// The MONET telescope (FB_MonetTelescopeControl) on mock axes, scanned in the MONETS MAIN order (telescope first, then
// the axes). One Scan() is one PLC scan. The scenario tests own one rig each (VAR_INST of the test method) and call Scan()
// once per PLC cycle: the astronomical clock needs a real NT_GetTime round trip (up to about 5 s) before the telescope
// accepts a goto/slew/track, so a rig is not usable before ClockValid. Everything else counts scans, not time.
// Plan: BROTLib specs/plans/2026-10-21-telescope-state-machine-unification.md (D1, step 1).
{attribute 'enable_dynamic_creation'}
FUNCTION_BLOCK FB_MonetRig
VAR
	fbComm			: FB_LogRecordingComm;	// #287: the log of the rig can be watched (fbComm.sWatch, nWatchHits)
	fbElev			: FB_ElevationMock(comm := fbComm);
	fbAzim			: FB_AzimuthMock(comm := fbComm);
	fbDero			: FB_DerotatorMock(comm := fbComm);
	fbFocus			: FB_FocusMock(comm := fbComm);
	fbCovers		: FB_CoversMock(comm := fbComm);	// a HalfBROT.FB_CoverControl subclass, its FB_Init takes comm
	stCoverOut		: HalfBROT.ST_CoverOut;	// the process outputs of the covers and the focus block (HalfBROT 0.14.0: VAR_IN_OUT stOut); the mocks do not use them
	stFocusOut		: HalfBROT.ST_FocusOut;
	fbBrakeHyd		: FB_BrakeHydraulicsMock;
	fbPointing		: FB_PointingModelForward(AOFF := 0.0, BNP := 0.0, AN_A := 0.0, AE_A := 0.0, NPAE := 0.0, EOFF := 0.0, AN_E := 0.0, AE_E := 0.0, TF := 0.0);	// zero coefficients
	fbPointingInv	: FB_PointingModelInversion(fbPointing := fbPointing);
	fbTel			: FB_MonetTelescopeControl(comm := fbComm);
	fbWatchdog		: FB_MonetMqttWatchdog(comm := fbComm);	// for MonetSafeState_Tests (a method VAR_INST cannot refer to a sibling in its init list)
	nScans			: UDINT;
	bManual			: BOOL;	// MAIN calls SuspendAutomatic instead of the body while the cabinet selector is on manual
	nTimeDivisor	: UDINT := 1;	// the time seam of the telescope under test (SetTimeDivisor)
	bEstopIn		: BOOL;	// SafetyHandling.estop
	bSafetyIn		: BOOL;	// SafetyHandling.error
	bMainReadyIn	: BOOL := TRUE;	// PowerMonitoring.phaseOK (MAIN: bMainReady := ready)
	stMotion		: BROTLib.ST_MotionConfig;	// stMotion of the telescope under test (SetMotion), default = the struct defaults (#24 step 2c)
	fElevationMoveVelocityIn	: LREAL := 5.0;	// the deprecated alias input (SetElevationMoveVelocity), default = its old default; MONETS MAIN passes 3.0
END_VAR
VAR CONSTANT
	telescopeConfig	: ST_TelescopeConfig := (longitude := 20.810808, latitude := -32.375823, altitude := 1798.0,
											 azimuthPark := 175, elevationPark := 60, derotatorPark := 0, focusPark := 36.0,
											 azimuthHome := 175, elevationHome := 40, derotatorHome := 0,
											 name := 'MONET/S', diameter := 1.2, cabinet := 'Beckhoff', manufacturer := 'test',
											 mountOptions := 'ALT-AZ', mount := 'ALT_AZ');
END_VAR

// scans a homing takes on the three mock axes (default 3): a test that wants to act while the axes are homing makes it longer
METHOD SetHomeScans
VAR_INPUT
	nScans	: UINT;
END_VAR
fbElev.nMockHomeScans := nScans;
fbAzim.nMockHomeScans := nScans;
fbDero.nMockHomeScans := nScans;
END_METHOD

// scans a move takes on the three mock axes (default 60)
METHOD SetMoveScans
VAR_INPUT
	nScans	: UINT;
END_VAR
fbElev.nMockMoveScans := nScans;
fbAzim.nMockMoveScans := nScans;
fbDero.nMockMoveScans := nScans;
END_METHOD

// 2026-11-11: TRUE = a move of the elevation/azimuth mock ends at the target of its start (MC_MoveAbsolute), not at the
// target of the scan it ends in (default FALSE, the model of the older tests)
METHOD SetMoveLatchesTarget
VAR_INPUT
	bValue	: BOOL;
END_VAR
fbElev.bMockLatchTarget := bValue;
fbAzim.bMockLatchTarget := bValue;
fbDero.bMockLatchTarget := bValue;
END_METHOD

// #267: the encoder of each mock axis lags its NC set position by this much (deg, ActualPosition = SetPosition - value), like the
// 1-3 mdeg of MONET/N at the end of a move; 0 (default) = ActualPosition and SetPosition are the same
METHOD SetFollowingError
VAR_INPUT
	fElevation	: LREAL;
	fAzimuth	: LREAL;
	fDerotator	: LREAL;
END_VAR
fbElev.fMockFollowingError := fElevation;
fbAzim.fMockFollowingError := fAzimuth;
fbDero.fMockFollowingError := fDerotator;
END_METHOD

// scans an MC_Stop takes on the three mock axes (default 3); a very large value is an axis that never reports standstill
METHOD SetStopScans
VAR_INPUT
	nScans	: UINT;
END_VAR
fbElev.nMockStopScans := nScans;
fbAzim.nMockStopScans := nScans;
fbDero.nMockStopScans := nScans;
END_METHOD

// divides every long timeout of the telescope (600 s, 2 min, 12 h) by nValue, for this rig only (1 = real times)
METHOD SetTimeDivisor
VAR_INPUT
	nValue	: UDINT;
END_VAR
nTimeDivisor := nValue;
fbTel.nTimeDivisor := nValue;	// also in manual, where the body (and its input list) is not called
END_METHOD

METHOD Scan
IF bManual THEN
	fbTel.SuspendAutomatic(bEstopIn := bEstopIn, bSafetyErrorIn := bSafetyIn, bMainReadyIn := bMainReadyIn);
ELSE
	fbTel(
		telescopeConfig := telescopeConfig,
		fbCovers := fbCovers,
		fbBrake := fbBrakeHyd,
		fbHydraulics := fbBrakeHyd,
		fbFocus := fbFocus,
		fbElevation := fbElev,
		fbAzimuth := fbAzim,
		fbDerotator := fbDero,
		fbPointing := fbPointing,
		fbPointingInverse := fbPointingInv,
		bEstopTriggered := bEstopIn,
		bSafetyError := bSafetyIn,
		bMainReady := bMainReadyIn,
		stMotion := stMotion,
		fElevationMoveVelocity := fElevationMoveVelocityIn,
		nTimeDivisor := nTimeDivisor);
END_IF
fbCovers(stOut := stCoverOut);	// after the telescope, as MAIN calls CoverControl(); only the travel model (SetCoverTravelScans) runs in it
fbElev(fbCovers := fbCovers, fbBrake := fbBrakeHyd);
fbAzim(bBrakeOpen := fbBrakeHyd.BrakeOpen, bMockBrakeGate := TRUE);	// #277: the azimuth enable needs the shared brake, as in HalfBROT
fbDero();
fbFocus(stOut := stFocusOut);
fbBrakeHyd();	// last: a close of this scan wins over the elevation's opening request (#272)
nScans := nScans + 1;
END_METHOD

PROPERTY ClockValid : BOOL
GET
ClockValid := fbTel.fbTime.bValid;
END_GET
END_PROPERTY

PROPERTY Online : BOOL
GET
Online := fbTel.ReadyState = 1.0;
END_GET
END_PROPERTY

// #287: the log messages of the rig that contained the text of WatchLog since that call
PROPERTY LogHits : INT
GET
LogHits := fbComm.nWatchHits;
END_GET
END_PROPERTY

// #287: count every log message of the rig that contains sText (LogHits), from now on
METHOD WatchLog
VAR_INPUT
	sText	: STRING(80);
END_VAR
fbComm.sWatch := sText;
fbComm.Clear();
END_METHOD

// stMotion of the telescope under test (#24 step 2c), handed to it from the next Scan() on; the default is the struct defaults
METHOD SetMotion
VAR_INPUT
	stValue	: BROTLib.ST_MotionConfig;
END_VAR
stMotion := stValue;
END_METHOD

// the deprecated alias input fElevationMoveVelocity of the telescope (#24 D2); 5.0 (default) = not used, MONETS MAIN passes 3.0
METHOD SetElevationMoveVelocity
VAR_INPUT
	fValue	: LREAL;
END_VAR
fElevationMoveVelocityIn := fValue;
END_METHOD

// the cabinet selector: TRUE = manual (the telescope body is not called, SuspendAutomatic is)
METHOD SetManual
VAR_INPUT
	bValue	: BOOL;
END_VAR
bManual := bValue;
END_METHOD

// scans a full open or close of the mock covers takes (default 0: at once); > 0 lets a test press the E-stop during a cover run
METHOD SetCoverTravelScans
VAR_INPUT
	nScans	: UINT;
END_VAR
fbCovers.nMockTravelScans := nScans;
END_METHOD

// the E-stop input of the telescope
METHOD SetEstop
VAR_INPUT
	bValue	: BOOL;
END_VAR
bEstopIn := bValue;
END_METHOD

// the safety error input of the telescope (SafetyHandling.error, #155)
METHOD SetSafetyError
VAR_INPUT
	bValue	: BOOL;
END_VAR
bSafetyIn := bValue;
END_METHOD

// writes the slew flag of the telescope directly (an ADS write); the methods reject a move before it is set while the clock is invalid
METHOD SetSlewFlag
fbTel.bSlew := TRUE;
END_METHOD

// #24 step 5: the slew input of the telescope as a level (an ADS write or a Visu button held or released); the telescope never
// writes it, its rising edge is the command
METHOD SetSlewInput
VAR_INPUT
	bValue	: BOOL;
END_VAR
fbTel.bSlew := bValue;
END_METHOD

// #24 step 5: the target inputs a slew input uses (what the Visu writes before the button: fAzimuth, fElevation)
METHOD SetSlewTargetInput
VAR_INPUT
	fAzimuth	: LREAL;
	fAltitude	: LREAL;
END_VAR
fbTel.fAzimuth := fAzimuth;
fbTel.fElevation := fAltitude;
END_METHOD

// the power input of the telescope (bMainReady, MAIN: PowerMonitoring.phaseOK); FALSE = power failure. Default TRUE.
METHOD SetMainReady
VAR_INPUT
	bValue	: BOOL;
END_VAR
bMainReadyIn := bValue;
END_METHOD

// the pendant jog button for the elevation (up)
METHOD JogElevation
VAR_INPUT
	bValue	: BOOL;
END_VAR
fbElev.MovePos := bValue;
END_METHOD

METHOD InjectElevationError
VAR_INPUT
	nId	: UDINT;
END_VAR
fbElev.InjectError(nId);
END_METHOD

// The elevation enable drops outside the telescope control (the ADS write of MONET/N run B, #277).
METHOD DisableElevation
fbElev.Enable := FALSE;
END_METHOD

METHOD InjectAzimuthError
VAR_INPUT
	nId	: UDINT;
END_VAR
fbAzim.InjectError(nId);
END_METHOD

METHOD InjectFocusError
VAR_INPUT
	nId	: UDINT;
END_VAR
fbFocus.InjectError(nId);
END_METHOD

METHOD InjectDerotatorError
VAR_INPUT
	nId	: UDINT;
END_VAR
fbDero.InjectError(nId);
END_METHOD

METHOD SetAzimuthPowerLost
VAR_INPUT
	bLost	: BOOL;
END_VAR
fbAzim.SetPowerLost(bLost);
END_METHOD

// #251: write the RA/Dec inputs of the telescope directly, like the Visu binding or an ADS client (not through Track()). A nested input cannot be written from a test (rig.fbTel.x).
METHOD SetTargetDirect
VAR_INPUT
	fRa		: LREAL;
	fDec	: LREAL;
END_VAR
fbTel.fRightAscension := fRa;
fbTel.fDeclination := fDec;
END_METHOD

// #251: the derotator guard of the retarget blend (default 0.005 deg)
METHOD SetRetargetDerotatorMax
VAR_INPUT
	fValue	: LREAL;
END_VAR
fbTel.fRetargetDerotatorMax := fValue;
END_METHOD

// BROTLib#167: bFeedFromPosition of the telescope
METHOD SetFeedFromPosition
VAR_INPUT
	bValue	: BOOL;
END_VAR
fbTel.bFeedFromPosition := bValue;
END_METHOD

END_FUNCTION_BLOCK

(* stored: Version 1.1.0.1, ProductVersion 3.1.4024.15
   POU FB_MonetRig: Id {60e92a7a-02cd-4e48-8d20-abdb7dc0369f}, SpecialFunc None
   Method SetHomeScans: Id {8a18ef85-bb7c-4844-b14a-04199381c5b4}
   Method SetMoveScans: Id {65c9910e-1c65-4968-95a1-8c415702ba7d}
   Method SetMoveLatchesTarget: Id {6bd8caef-7020-4a79-98db-931b4c9b80ef}
   Method SetFollowingError: Id {77b0b675-340b-4379-8d7a-5ee7568305c9}
   Method SetStopScans: Id {d676b49d-f214-4b42-a004-df2964ff2f3e}
   Method SetTimeDivisor: Id {ebf41625-64f0-473d-96e0-0430a16c873f}
   Method Scan: Id {121ba66a-36ff-4009-9705-7efd4e908f1b}
   Property ClockValid: Id {3076ff3c-98ad-4dc0-97fb-ed4821c83c33}
   Get Get: Id {bc2a52f7-905d-4428-b9c8-29b6c1c1c00d}
   Property Online: Id {d88bbb8d-d30d-4985-b3f0-0b0b689944f1}
   Get Get: Id {fa836018-c28d-4e5d-becc-884b5bb557c9}
   Property LogHits: Id {42f1f42d-ff27-434c-8907-925c6dd494b4}
   Get Get: Id {ecc727e9-b181-4cc8-8945-00961633fa5a}
   Method WatchLog: Id {46326d1d-eeb3-445f-8073-898474c30993}
   Method SetMotion: Id {a8848ecf-4ba6-4d7f-95e4-4a32a59465d5}
   Method SetElevationMoveVelocity: Id {62399cab-459e-47e6-bff3-27d83498d3ec}
   Method SetManual: Id {7367e2f8-5967-47be-afd4-0d6ea17370fa}
   Method SetCoverTravelScans: Id {44131a3b-7ab9-4087-a9e2-27fc7d8d14c2}
   Method SetEstop: Id {f76d3ba5-df1c-4f8b-afcc-6f56a0d9547e}
   Method SetSafetyError: Id {a8622214-e2e0-447a-aac1-516f64995742}
   Method SetSlewFlag: Id {acff02fe-462d-4119-ba0f-3270ddb40627}
   Method SetSlewInput: Id {7befd08b-db5e-4357-97aa-6eb3458cdf4a}
   Method SetSlewTargetInput: Id {26be7ad4-8976-4b6a-86eb-973975e56a4f}
   Method SetMainReady: Id {83eaab32-d382-48b6-babc-99dec72544d2}
   Method JogElevation: Id {99a17950-974a-44cd-b2a3-f86293f3314d}
   Method InjectElevationError: Id {4c2738fe-bd1d-4e40-8884-048309dc8e4b}
   Method DisableElevation: Id {157508e2-dd45-48fd-8139-697da48b8a16}
   Method InjectAzimuthError: Id {5857afe2-6b7e-47e4-849f-b3e7bfb14aca}
   Method InjectFocusError: Id {f0de967d-0d68-41a5-ad3e-328e6c9af1d2}
   Method InjectDerotatorError: Id {b1bf17dc-df53-46f0-a8d3-000210700a06}
   Method SetAzimuthPowerLost: Id {90980f09-40a4-4fe6-bdab-e7ed198b3590}
   Method SetTargetDirect: Id {6ca861a5-2b2b-43f7-84ea-69efe59eab8a}
   Method SetRetargetDerotatorMax: Id {447a6f6b-55f7-4c2a-b1bf-373b727d9a02}
   Method SetFeedFromPosition: Id {05e47d2a-3fd2-4173-8991-5a2fb09bc14d} *)
